(* CODESYS project Live_Visu.vis.xml

Project tree, tasks and I/O mapping:
  visualisation Live_Visu
*)

// /Live_Visu
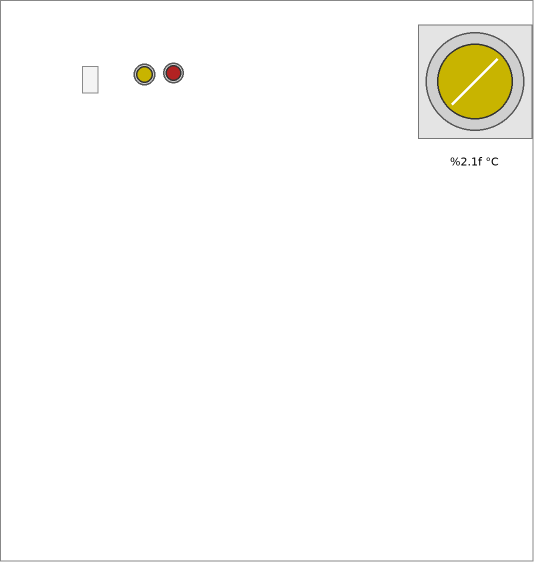
VISUALIZATION Live_Visu  // 534x562
    Polygon (13,14) (261,7) (373,51) (69,61)
    Polygon (77,61) (367,52) (367,75) (76,90)
    Polygon (69,61) (77,61) (77,89) (73,91) (66,89)
    Polygon (13,13) (68,61) (67,91) (13,43)
    Polygon (367,51) (377,51) (376,73) (367,74)
    Potentiometer360 (418,24 114x115), variable: Glob_Var.TempSet, style: Potentiometer-Potentiometer360-Yellow, scale format: %.0f, scale 3..13
        p2431819421: Outside
        p518627256: °C
    Rectangle (426,145 97x34), "%2.1f °C", text variable: Glob_Var.TempActual
    Lamp1 (132,62 25x25), variable: Glob_Var.Compressor, style: Lamp-Lamp1-Yellow
    Lamp1 (161,61 25x24), variable: Glob_Var.Signal, style: Lamp-Lamp1-Red
    Group (66,75 301x465)
        Polygon (3,17) (301,0) (292,422) (5,465) (2,464)
        Group (0,30 33x119)
            Polygon (2,0) (18,1) (22,11) (28,29) (32,46) (33,67) (31,84) (27,97) (22,108) (16,119) (3,117) (15,97) (18,84) (20,70) (20,48) (15,27) (9,14)
            Polygon (3,0) (0,1) (0,5) (3,8) (5,12) (8,16) (10,20) (12,26) (13,31) (16,40) (17,46) (18,54) (18,62) (18,72) (16,80) (14,89) (11,97) (7,106) (2,117) (4,118) (9,107) (13,100) (17,90) (19,80) (21,69) (21,62) (20,48) (17,36) (15,27) (10,14) (7,7)
    Polygon (13,45) (66,92) (69,539) (12,412)
    Group (65,78 299x482), invisible if: NOT Glob_Var.DoorOpen
        Polygon (1,17) (299,0) (290,422) (3,465) (0,464)
        Group (21,0 278x482)
            Polygon (1,34) (278,0) (270,421) (3,482) (0,481)
            Group (1,69 33x119)
                Polygon (2,0) (18,1) (22,11) (28,29) (32,46) (33,67) (31,84) (27,97) (22,108) (16,119) (3,117) (15,97) (18,84) (20,70) (20,48) (15,27) (9,14)
                Polygon (3,0) (0,1) (0,5) (3,8) (5,12) (8,16) (10,20) (12,26) (13,31) (16,40) (17,46) (18,54) (18,62) (18,72) (16,80) (14,89) (11,97) (7,106) (2,117) (4,118) (9,107) (13,100) (17,90) (19,80) (21,69) (21,62) (20,48) (17,36) (15,27) (10,14) (7,7)
    RockerSwitch (82,66 16x27), variable: Glob_Var.DoorOpen, behaviour: TOGGLE, style: Switch-RockerSwitch-Gray
END_VISUALIZATION
